Fanuc KAREL source: kc00028.KL

-- PROVISIONAL review KL for V1013-1; original PC SHA256 69dbab4b27d0635452ab7432255cebab01ed06bda0a8ecbca3f5a132d212365b
-- Incomplete behavior may be omitted. Consult companion uncertainty JSON. Do not deploy.
PROGRAM KC00028
%NOLOCKGROUP
BEGIN
  -- UNRESOLVED_PC offsets 5-93; opcodes 27,22,1C,22,1C,22,1C,22,1C,22,22,22,22,1C,22,31
  -- UNRESOLVED_PC offsets 98-102; opcodes 7F
END KC00028
